// TIA Portal V18 export
DATA_BLOCK "TEST_OPC_UA"   // DB3
{ S7_Optimized_Access := 'TRUE' }
// stored: MemoryReserve 100
   VAR
      Static_1TESTGIT : Real := 1.0;
      TEMP_1 : Real := 2.0;
      TEMP_2 : Real := 3.0;
      TEMP_3 : Real := 4.0;
      TEMP_4 : Real := 5.0;
      TEMP_5 : Real := 6.0;
      TEMP_6 : Real := 7.0;
   END_VAR
BEGIN
END_DATA_BLOCK
